(* Logix 5000 project; controller TFF vendor 1 type 14 code 107 rev 34.11; software revision 34.03; part 18 of 36 *)
(* tags used below, declared in another part *)
   AlarmControl : AlarmControl;   // Alarm Control
   ControlLoop : ControlLoop[20];   // Control Loop Array
   ControlLoop_PCV001_5ms : ALIAS FOR ControlLoop[4];   // PCV001 Control Loop
   ControlLoop_PCV101 : ALIAS FOR ControlLoop[5];   // PCV101 Control Loop
   ControlLoop_PCV101_5ms : ALIAS FOR ControlLoop[6];   // PCV101 Control Loop
   ControlLoop_PCV101Alarm : ALIAS FOR AlarmDeviation[5];   // PCV101 Control Loop Deviation Alarm
   CPU_Scanning : BOOL;   // System Scanning Flag
   DigitalOutput : BOOL[256];   // Digital Output Array these bits are sent to output cards.
   FI101 : ALIAS FOR AnalogPoint[2];   // Filtrate Flow
   FirstScanComplete : BOOL;   // First Scan Complete Flag
   LI001 : ALIAS FOR AnalogPoint[44];   // Feed Bag Volume
   Membrane_Data : Membrane_Data;   // Membrane Data
   Options : Options;   // Options List
   PCV001 : ALIAS FOR AnalogPoint[3];   // Retentate Pressure Control Valve Position
   PCV101 : ALIAS FOR AnalogPoint[4];   // Filtrate Pressure Control Valve Position
   PCV101_AO : ALIAS FOR AnalogOutput[1];   // FiltratePressure Control Valve Setpoint
   PCV101_Control : PCV_Control;   // PCV101 Control UDT
   Phase0 : ALIAS FOR Phase[0];   // Phase 0
   PLCFault : FaultRecordType;   // PLC Major Fault Record
   Rack_Murr_Node1_TF2S : IO_Station;   // Status of Node 1 TF2S
   Rack_Murr_Node1_TF3S : IO_Station;   // Status of Node 1 TF3S
   Rack_Murr_Node6_IND331_WI001 : IO_Station;   // Status of Node 6 IND331 WI001
   Rack_Murr_Node7_IND131_WI101 : IO_Station;   // Status of Node 7 IND131 WI101
   RawAnalogInputArray : INT[50];   // Array of analog input raw
   ScaleFiltering : ScaleFiltering;   // Data for Scale Filtering
   SIC001 : ALIAS FOR Drive[1];   // Feed Pump
   SIC002 : ALIAS FOR Drive[2];   // Transfer Pump
   SysControl : SysControl;   // General system status and command
   ThisSystem : SystemType;
   TMP : ALIAS FOR AnalogPoint[41];   // Trans-membrane Pressure
   Valve : Valve[100];   // Valve Array
   ValveControl : ValveControl;   // Valve Control
   WI001 : ALIAS FOR AnalogPoint[15];   // Feed Bag Weight
   WI001Alarm : ALIAS FOR AlarmAnalog[15];   // Feed Bag Weight Alarm
   WI101 : ALIAS FOR AnalogPoint[0];   // Filtrate Weight
   WI101Alarm : ALIAS FOR AlarmAnalog[0];   // Filtrate Weight Alarm
   WI102 : ALIAS FOR AnalogPoint[1];   // Customer Filtrate Weight
   WI102Alarm : ALIAS FOR AlarmAnalog[1];   // Customer Filtrate Weight Alarm
   YA10 : ALIAS FOR DigitalPoint[59];   // PLC Program Major Fault
(* MainProgram5ms, continued *)

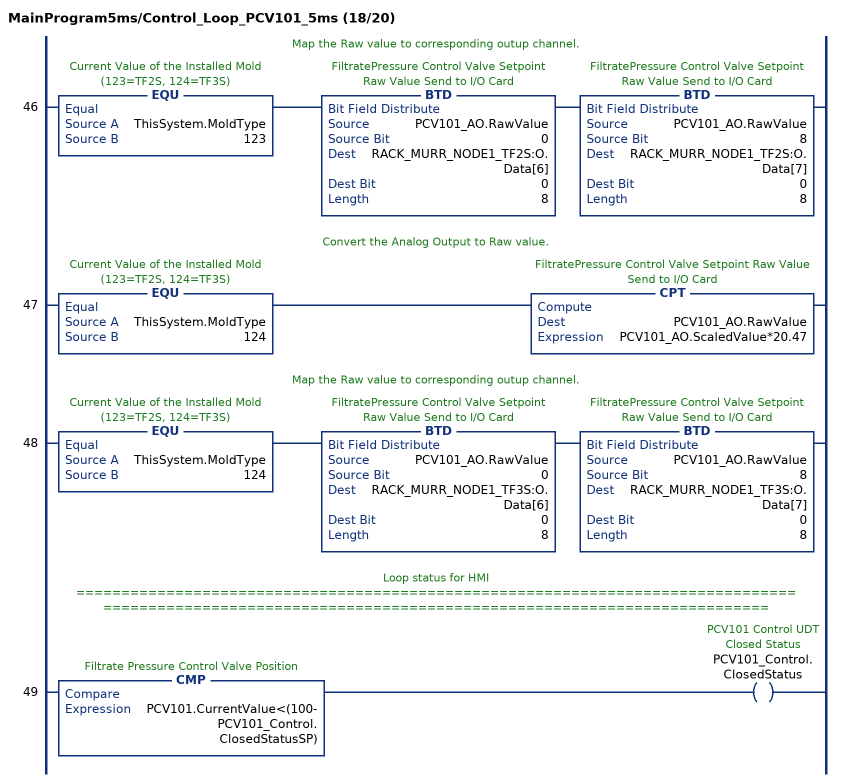
   // Map the Raw value to corresponding outup channel.
   46: EQU(ThisSystem.MoldType,123)BTD(PCV101_AO.RawValue,0,RACK_MURR_NODE1_TF2S:O.Data[6],0,8)BTD(PCV101_AO.RawValue,8,RACK_MURR_NODE1_TF2S:O.Data[7],0,8);
   // Convert the Analog Output to Raw value.
   47: EQU(ThisSystem.MoldType,124)CPT(PCV101_AO.RawValue,PCV101_AO.ScaledValue*20.47);
   // Map the Raw value to corresponding outup channel.
   48: EQU(ThisSystem.MoldType,124)BTD(PCV101_AO.RawValue,0,RACK_MURR_NODE1_TF3S:O.Data[6],0,8)BTD(PCV101_AO.RawValue,8,RACK_MURR_NODE1_TF3S:O.Data[7],0,8);
   // Loop status for HMI
   // ==========================================================================================================================================================
   49: CMP(PCV101.CurrentValue<(100-PCV101_Control.ClosedStatusSP))OTE(PCV101_Control.ClosedStatus);
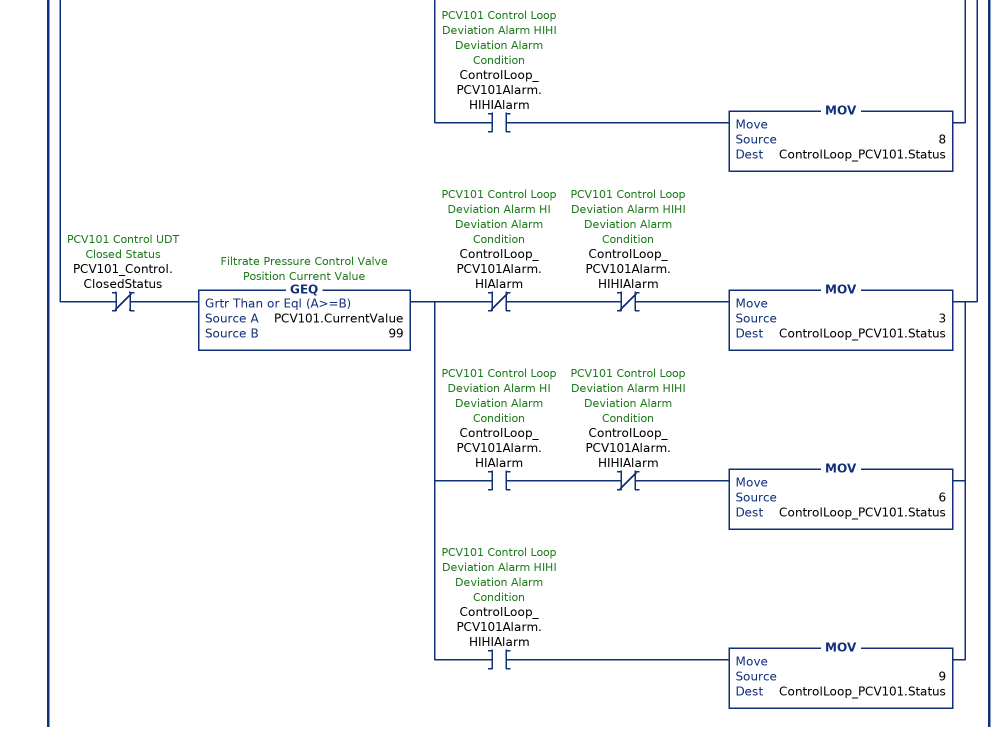
   // ControlLoop Status : 1 = PCV Close
   // ControlLoop Status : 2 = PCV Open
   // ControlLoop Status : 3 = PCV Full Open
   // ControlLoop Status : 4 = PCV Close and Non Critical alam
   // ControlLoop Status : 5 = PCV Open and Non Critical alam
   // ControlLoop Status : 6 = PCV Full Open and Non Critical alam
   // ControlLoop Status : 7 = PCV Close and Critical alam
   // ControlLoop Status : 8 = PCV Open and Critical alam
   // ControlLoop Status : 9 = PCV Full Open and Critical alam
   50: [XIC(PCV101_Control.ClosedStatus) [XIO(ControlLoop_PCV101Alarm.HIAlarm) XIO(ControlLoop_PCV101Alarm.HIHIAlarm) MOV(1,ControlLoop_PCV101.Status) ,XIC(ControlLoop_PCV101Alarm.HIAlarm) XIO(ControlLoop_PCV101Alarm.HIHIAlarm) MOV(4,ControlLoop_PCV101.Status) ,XIC(ControlLoop_PCV101Alarm.HIHIAlarm) MOV(7,ControlLoop_PCV101.Status) ] ,XIO(PCV101_Control.ClosedStatus) LES(PCV101.CurrentValue,99) [XIO(ControlLoop_PCV101Alarm.HIAlarm) XIO(ControlLoop_PCV101Alarm.HIHIAlarm) MOV(2,ControlLoop_PCV101.Status) ,XIC(ControlLoop_PCV101Alarm.HIAlarm) XIO(ControlLoop_PCV101Alarm.HIHIAlarm) MOV(5,ControlLoop_PCV101.Status) ,XIC(ControlLoop_PCV101Alarm.HIHIAlarm) MOV(8,ControlLoop_PCV101.Status) ] ,XIO(PCV101_Control.ClosedStatus) GEQ(PCV101.CurrentValue,99) [XIO(ControlLoop_PCV101Alarm.HIAlarm) XIO(ControlLoop_PCV101Alarm.HIHIAlarm) MOV(3,ControlLoop_PCV101.Status) ,XIC(ControlLoop_PCV101Alarm.HIAlarm) XIO(ControlLoop_PCV101Alarm.HIHIAlarm) MOV(6,ControlLoop_PCV101.Status) ,XIC(ControlLoop_PCV101Alarm.HIHIAlarm) MOV(9,ControlLoop_PCV101.Status) ] ];
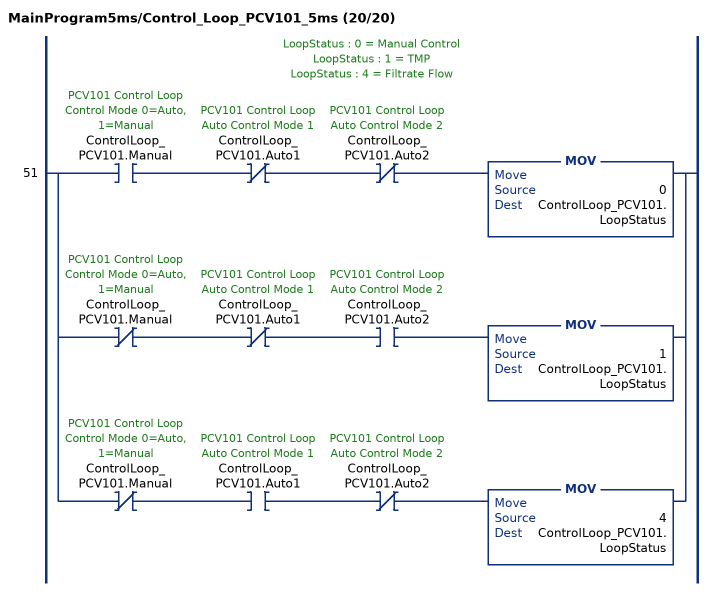
   // LoopStatus : 0 = Manual Control
   //  LoopStatus : 1 = TMP
   //  LoopStatus : 4 = Filtrate Flow
   51: [XIC(ControlLoop_PCV101.Manual) XIO(ControlLoop_PCV101.Auto1) XIO(ControlLoop_PCV101.Auto2) MOV(0,ControlLoop_PCV101.LoopStatus) ,XIO(ControlLoop_PCV101.Manual) XIO(ControlLoop_PCV101.Auto1) XIC(ControlLoop_PCV101.Auto2) MOV(1,ControlLoop_PCV101.LoopStatus) ,XIO(ControlLoop_PCV101.Manual) XIC(ControlLoop_PCV101.Auto1) XIO(ControlLoop_PCV101.Auto2) MOV(4,ControlLoop_PCV101.LoopStatus) ];
END_ROUTINE

ROUTINE FaultRoutine   (* ladder *)
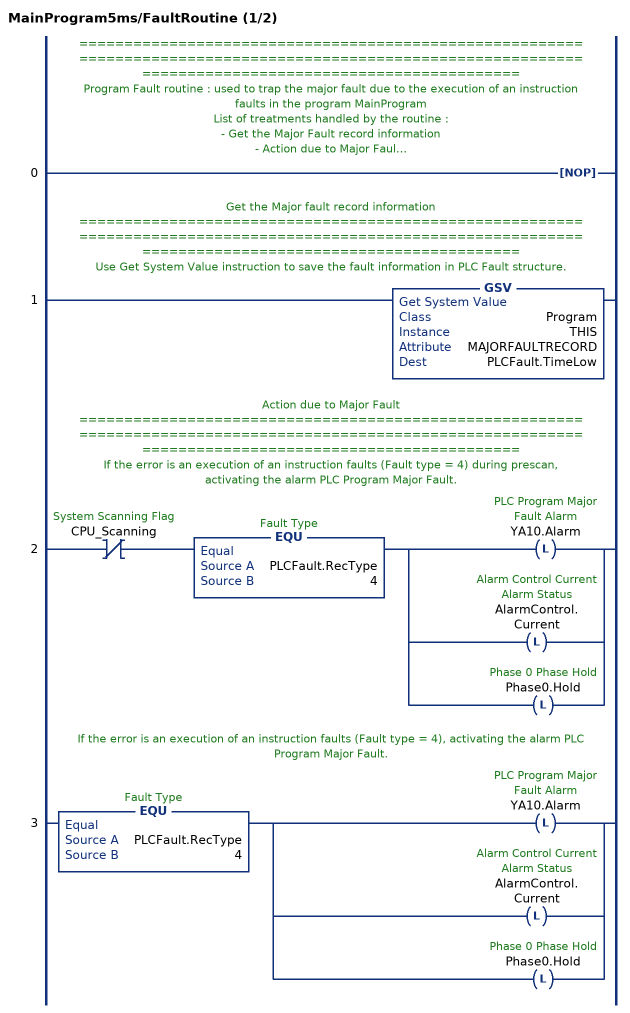
   // ==========================================================================================================================================================
   //                                                               Program Fault routine : used to trap the major fault due to the execution of an instruction faults in the program MainProgram
   //                                                     List of treatments handled by the routine :
   //                                                          - Get the Major Fault record information
   //                                                          - Action due to Major Fault
   //                                                     -----------------------------------------------------------------------------------------------------------------------------------------------------
   //                                                     History
   //                                                          2019-AUG-13 - Actemium - B. Roch - Initial version for Candidate Release 3.00.00.00.a
   // ==========================================================================================================================================================
   0: NOP();
   // Get the Major fault record information
   // ==========================================================================================================================================================
   // Use Get System Value instruction to save the fault information in PLC Fault structure.
   1: GSV(Program,THIS,MAJORFAULTRECORD,PLCFault.TimeLow);
   // Action due to Major Fault
   // ==========================================================================================================================================================
   // If the error is an execution of an instruction faults (Fault type = 4) during prescan, activating the alarm PLC Program Major Fault.
   2: XIO(CPU_Scanning)EQU(PLCFault.RecType,4)[OTL(YA10.Alarm) ,OTL(AlarmControl.Current) ,OTL(Phase0.Hold) ];
   // If the error is an execution of an instruction faults (Fault type = 4), activating the alarm PLC Program Major Fault.
   3: EQU(PLCFault.RecType,4)[OTL(YA10.Alarm) ,OTL(AlarmControl.Current) ,OTL(Phase0.Hold) ];
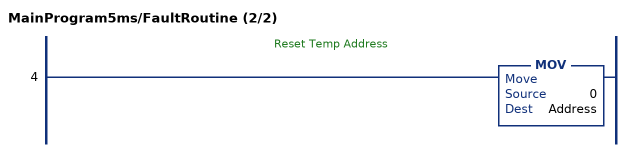
   // Reset Temp Address
   4: MOV(0,Address);
END_ROUTINE

ROUTINE Input_Analog_HighSpeed   (* ladder *)
// HighSpeed Analog Input Scaling
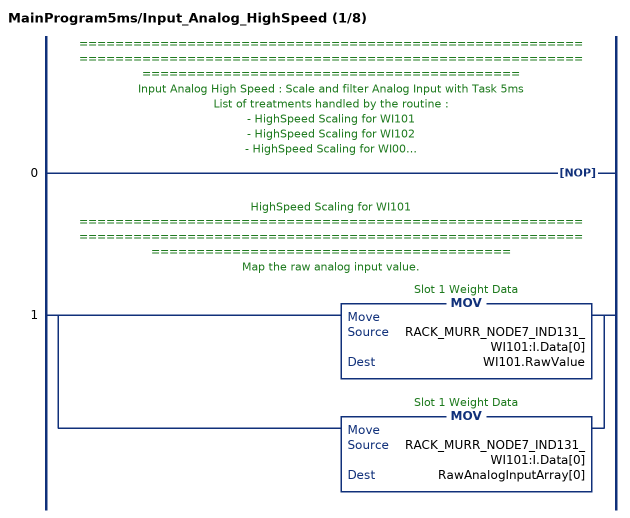
   // ==========================================================================================================================================================
   //                                                  Input Analog High Speed : Scale and filter Analog Input with Task 5ms
   //                                                     List of treatments handled by the routine :
   //                                                     - HighSpeed Scaling for WI101
   //                                                     - HighSpeed Scaling for WI102
   //                                                     - HighSpeed Scaling for WI001
   //                                                     - Scale Filtering processing
   //                                                     - Alarm Process Value Initialization
   //                                                     -----------------------------------------------------------------------------------------------------------------------------------------------------
   //                                                     History
   //                                                   2019-AUG-13 - Actemium - B. Roch - Initial version for Candidate Release 3.00.00.00.a                    		2019-SEP-11 - ACTEMIUM - Q. Spindler - Modifications for Candidate Release 3.00.00.00.c
   // 					- Change raw value for WI102 to 1
   // ==========================================================================================================================================================
   0: NOP();
   // HighSpeed Scaling for WI101
   // ========================================================================================================================================================
   // Map the raw analog input value.
   1: [MOV(RACK_MURR_NODE7_IND131_WI101:I.Data[0],WI101.RawValue) ,MOV(RACK_MURR_NODE7_IND131_WI101:I.Data[0],RawAnalogInputArray[0]) ];
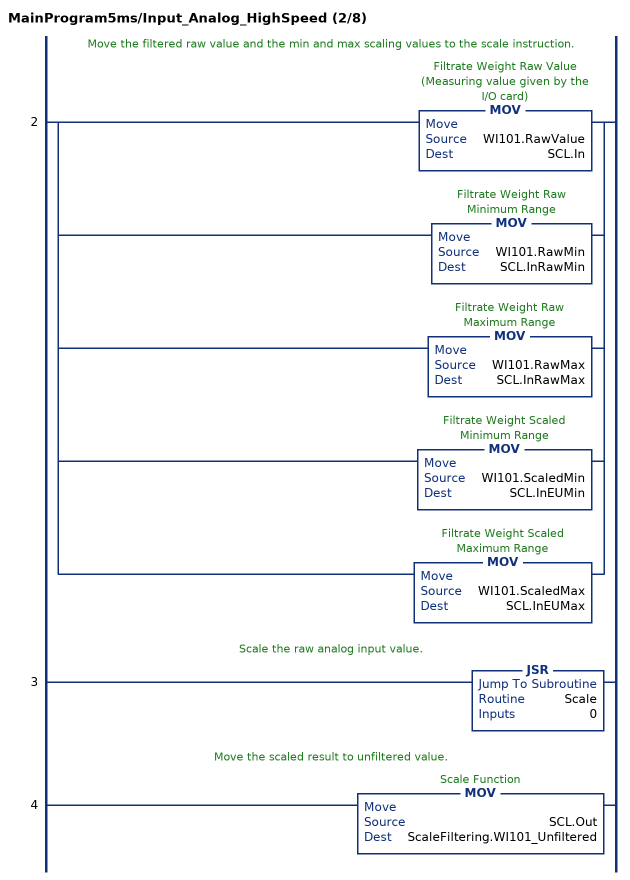
   // Move the filtered raw value and the min and max scaling values to the scale instruction.
   2: [MOV(WI101.RawValue,SCL.In) ,MOV(WI101.RawMin,SCL.InRawMin) ,MOV(WI101.RawMax,SCL.InRawMax) ,MOV(WI101.ScaledMin,SCL.InEUMin) ,MOV(WI101.ScaledMax,SCL.InEUMax) ];
   // Scale the raw analog input value.
   3: JSR(Scale,0);
   // Move the scaled result to unfiltered value.
   4: MOV(SCL.Out,ScaleFiltering.WI101_Unfiltered);
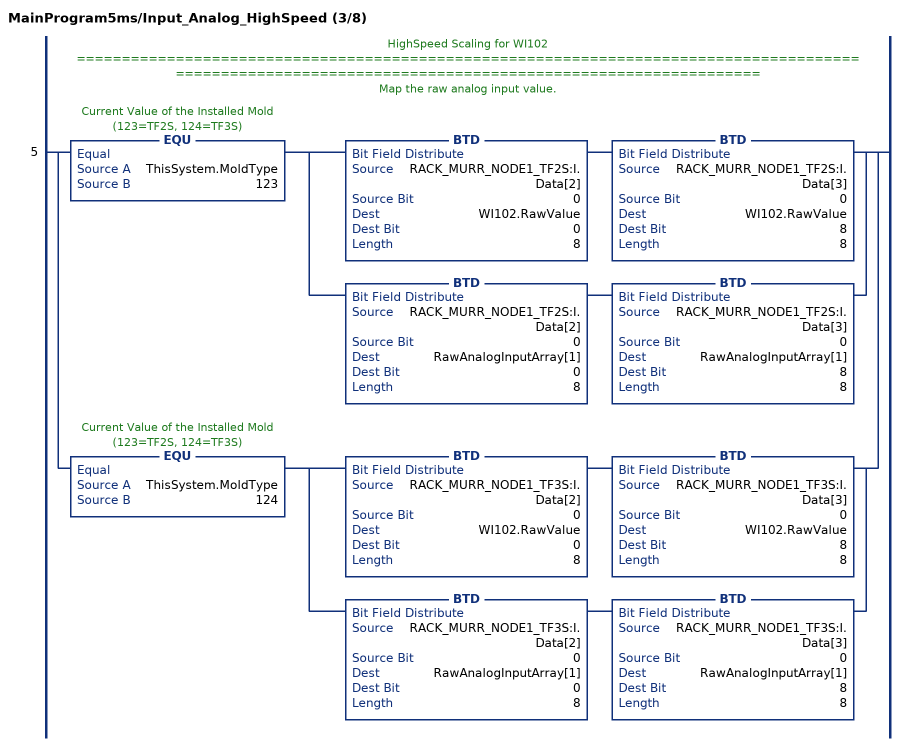
   // HighSpeed Scaling for WI102
   // ========================================================================================================================================================
   // Map the raw analog input value.
   5: [EQU(ThisSystem.MoldType,123) [BTD(RACK_MURR_NODE1_TF2S:I.Data[2],0,WI102.RawValue,0,8) BTD(RACK_MURR_NODE1_TF2S:I.Data[3],0,WI102.RawValue,8,8) ,BTD(RACK_MURR_NODE1_TF2S:I.Data[2],0,RawAnalogInputArray[1],0,8) BTD(RACK_MURR_NODE1_TF2S:I.Data[3],0,RawAnalogInputArray[1],8,8) ] ,EQU(ThisSystem.MoldType,124) [BTD(RACK_MURR_NODE1_TF3S:I.Data[2],0,WI102.RawValue,0,8) BTD(RACK_MURR_NODE1_TF3S:I.Data[3],0,WI102.RawValue,8,8) ,BTD(RACK_MURR_NODE1_TF3S:I.Data[2],0,RawAnalogInputArray[1],0,8) BTD(RACK_MURR_NODE1_TF3S:I.Data[3],0,RawAnalogInputArray[1],8,8) ] ];
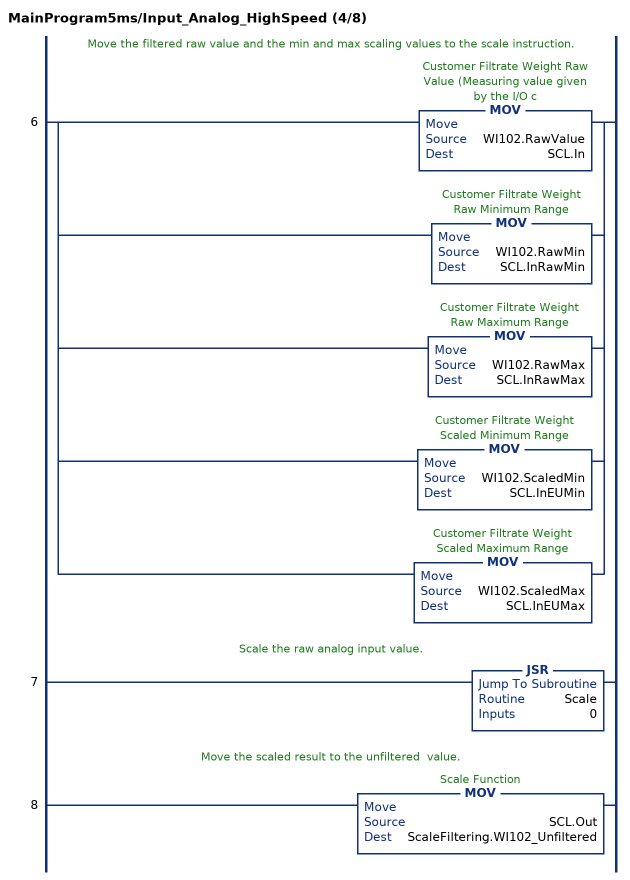
   // Move the filtered raw value and the min and max scaling values to the scale instruction.
   6: [MOV(WI102.RawValue,SCL.In) ,MOV(WI102.RawMin,SCL.InRawMin) ,MOV(WI102.RawMax,SCL.InRawMax) ,MOV(WI102.ScaledMin,SCL.InEUMin) ,MOV(WI102.ScaledMax,SCL.InEUMax) ];
   // Scale the raw analog input value.
   7: JSR(Scale,0);
   // Move the scaled result to the unfiltered  value.
   8: MOV(SCL.Out,ScaleFiltering.WI102_Unfiltered);
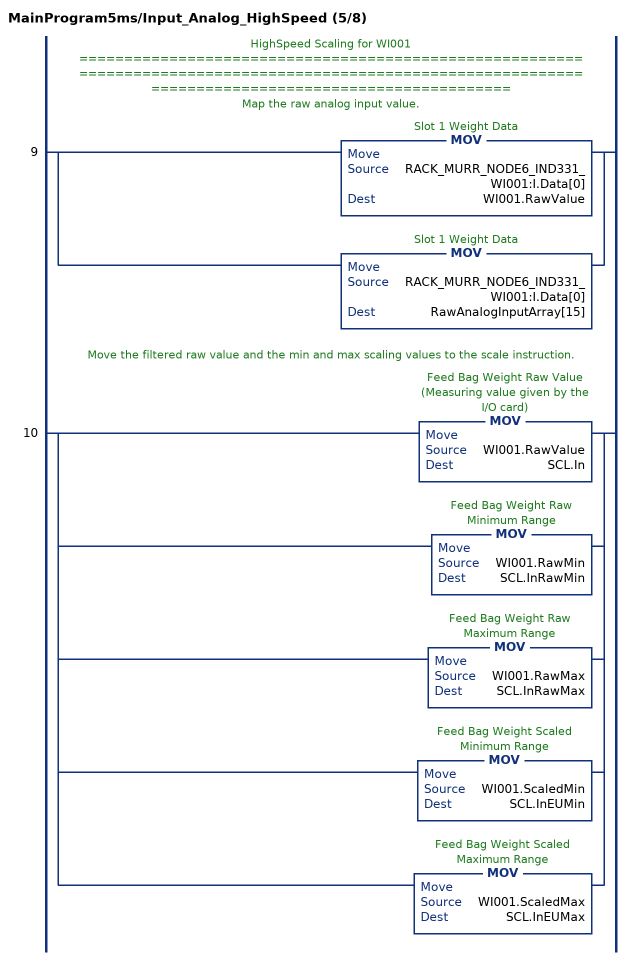
   // HighSpeed Scaling for WI001
   // ========================================================================================================================================================
   // Map the raw analog input value.
   9: [MOV(RACK_MURR_NODE6_IND331_WI001:I.Data[0],WI001.RawValue) ,MOV(RACK_MURR_NODE6_IND331_WI001:I.Data[0],RawAnalogInputArray[15]) ];
   // Move the filtered raw value and the min and max scaling values to the scale instruction.
   10: [MOV(WI001.RawValue,SCL.In) ,MOV(WI001.RawMin,SCL.InRawMin) ,MOV(WI001.RawMax,SCL.InRawMax) ,MOV(WI001.ScaledMin,SCL.InEUMin) ,MOV(WI001.ScaledMax,SCL.InEUMax) ];
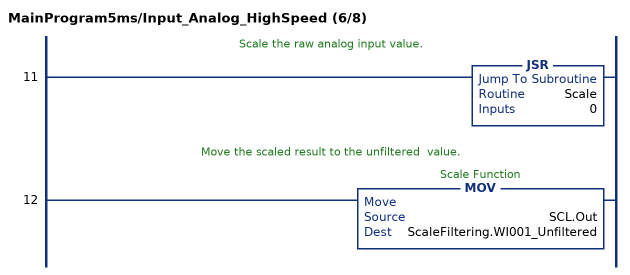
   // Scale the raw analog input value.
   11: JSR(Scale,0);
   // Move the scaled result to the unfiltered  value.
   12: MOV(SCL.Out,ScaleFiltering.WI001_Unfiltered);
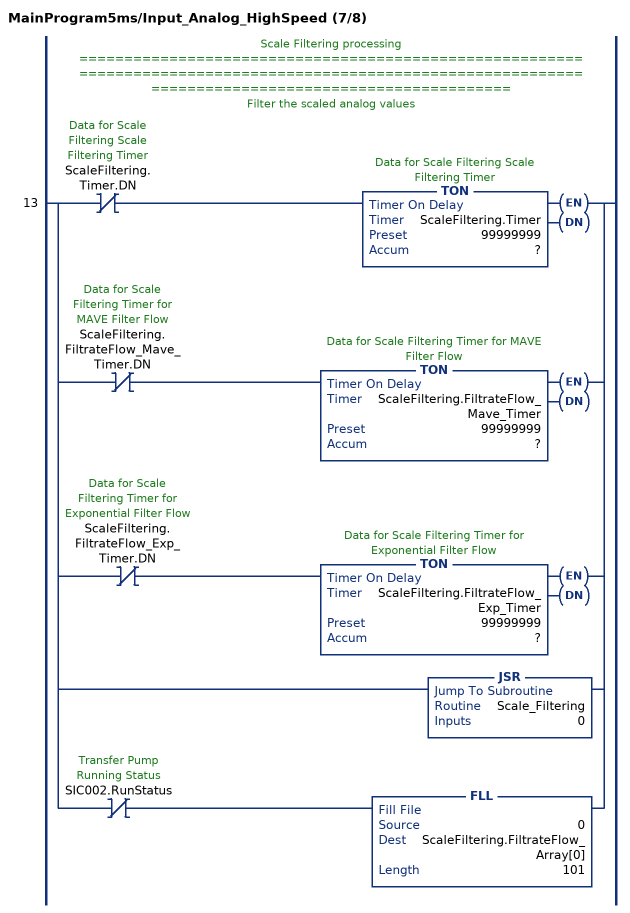
   // Scale Filtering processing
   // ========================================================================================================================================================
   // Filter the scaled analog values
   13: [XIO(ScaleFiltering.Timer.DN) TON(ScaleFiltering.Timer,?,?) ,XIO(ScaleFiltering.FiltrateFlow_Mave_Timer.DN) TON(ScaleFiltering.FiltrateFlow_Mave_Timer,?,?) ,XIO(ScaleFiltering.FiltrateFlow_Exp_Timer.DN) TON(ScaleFiltering.FiltrateFlow_Exp_Timer,?,?) ,JSR(Scale_Filtering,0) ,XIO(SIC002.RunStatus) FLL(0,ScaleFiltering.FiltrateFlow_Array[0],101) ];
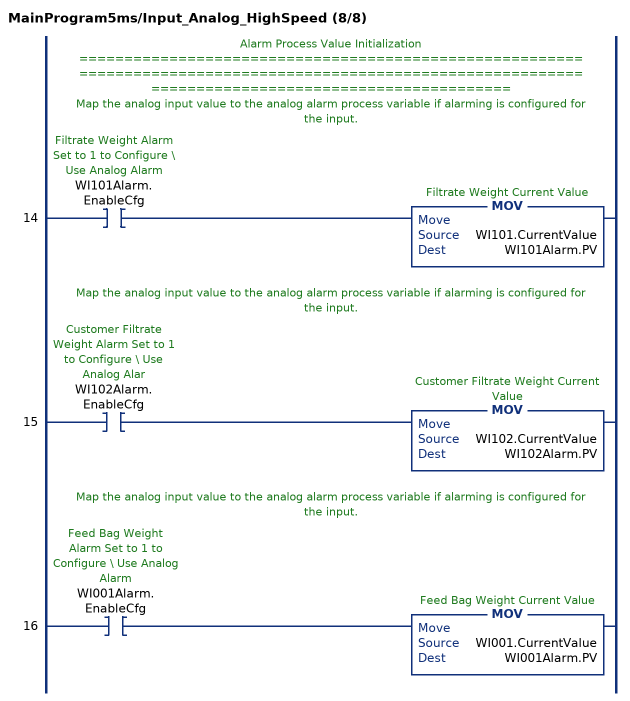
   // Alarm Process Value Initialization
   // ========================================================================================================================================================
   // Map the analog input value to the analog alarm process variable if alarming is configured for the input.
   14: XIC(WI101Alarm.EnableCfg)MOV(WI101.CurrentValue,WI101Alarm.PV);
   // Map the analog input value to the analog alarm process variable if alarming is configured for the input.
   15: XIC(WI102Alarm.EnableCfg)MOV(WI102.CurrentValue,WI102Alarm.PV);
   // Map the analog input value to the analog alarm process variable if alarming is configured for the input.
   16: XIC(WI001Alarm.EnableCfg)MOV(WI001.CurrentValue,WI001Alarm.PV);
END_ROUTINE

ROUTINE MainRoutine   (* ladder *)
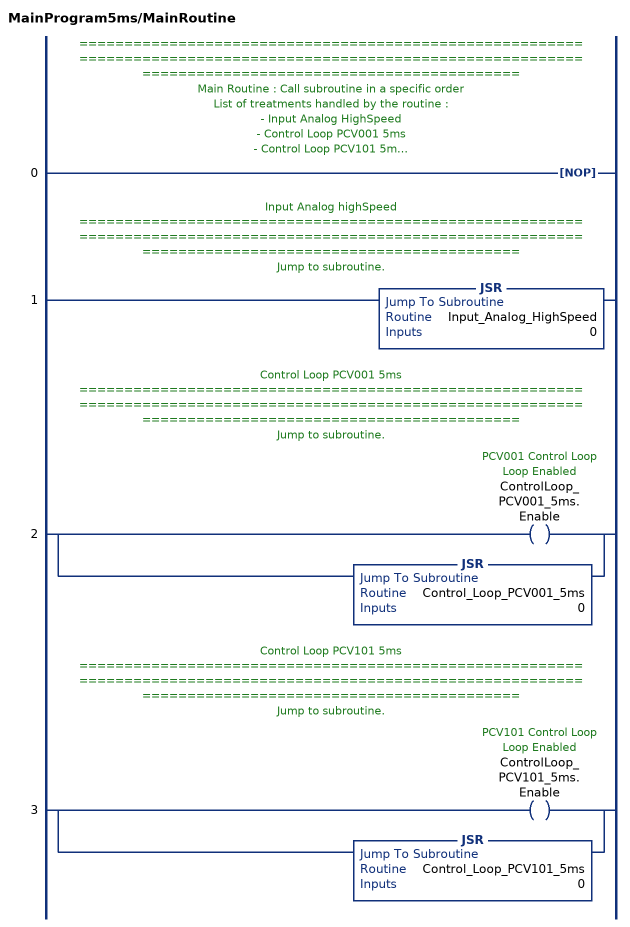
   // ==========================================================================================================================================================
   //                                                  Main Routine : Call subroutine in a specific order
   //                                                     List of treatments handled by the routine :
   //                                                - Input Analog HighSpeed
   //                                                - Control Loop PCV001 5ms
   //                                                - Control Loop PCV101 5ms
   //                                                     -----------------------------------------------------------------------------------------------------------------------------------------------------
   //                                                     History
   //                                                        2019-AUG-13 - Actemium - B. Roch - Initial version for Candidate Release 3.00.00.00.a
   // ==========================================================================================================================================================
   0: NOP();
   // Input Analog highSpeed
   // ==========================================================================================================================================================
   // Jump to subroutine.
   1: JSR(Input_Analog_HighSpeed,0);
   // Control Loop PCV001 5ms
   // ==========================================================================================================================================================
   // Jump to subroutine.
   2: [OTE(ControlLoop_PCV001_5ms.Enable) ,JSR(Control_Loop_PCV001_5ms,0) ];
   // Control Loop PCV101 5ms
   // ==========================================================================================================================================================
   // Jump to subroutine.
   3: [OTE(ControlLoop_PCV101_5ms.Enable) ,JSR(Control_Loop_PCV101_5ms,0) ];
END_ROUTINE

ROUTINE Scale   (* function block diagram *)
// Scale Routine
   SHEET 1
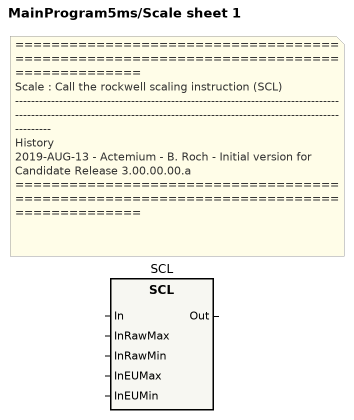
   // ======================================================================================
   // Scale : Call the rockwell scaling instruction (SCL)
   // ------------------------------------------------------------------------------------------------------------------------------------------------------------------
   // ---------
   // History
   //    2019-AUG-13 - Actemium - B. Roch - Initial version for Candidate Release 3.00.00.00.a
   // ======================================================================================
   SCL : SCL();   // unwired pins: In InRawMax InRawMin InEUMax InEUMin Out
END_ROUTINE

ROUTINE Scale_Filtering   (* structured text *)
   
   (* =======================================================================
   	Scale Filtering : calculations of Filtered value
   
   	List of treatments
   		- Initialize Volume
   		- WI001 Feed Bag Volume Calculation
   		- Moving Average Filtering for Filtrate Volume
   		- Moving Average Filtering for Filtrate Flow
   		- Exponential Filtering for Filtrate Volume
   		- Exponential Filtering for Filtrate Flow
   		- Analog Input processing
   
   -----------------------------------------------------------------------------------------------------------------------------------------------------
   	History
   		2019-AUG-13 - ACTEMIUM - B. Roch - Initial version for Candidate Release 3.00.00.00.a
   		2019-SEP-17 - ACTEMIUM - Q. Spindler - Modifications for Candidate Release 3.00.00.00.c
   					- Bypass CurrentValue calculation when in simulation mode
   					- Remove Initialize Values as they will be stored in CCPSettings
   =============================================================================================================================*)
   
   
   
   (* Initialize Volume
   =============================================================================================================================*)
   
   // Compute Volume values based on Unfiltered Weight and Density
   ScaleFiltering.FeedBagVolume := ScaleFiltering.WI001_Unfiltered / Membrane_Data.Density;
   ScaleFiltering.FiltrateVolume101 := ScaleFiltering.WI101_Unfiltered / Membrane_Data.Density;
   ScaleFiltering.FiltrateVolume102 := ScaleFiltering.WI102_Unfiltered / Membrane_Data.Density;
   
   
   //Check that the minimum sample rate have met
   If ScaleFiltering.Timer.ACC > ScaleFiltering.Sample_Rate Then
   
   (* WI001 Feed Bag Volume Calculation
   =============================================================================================================================*)
   
   		//Compute the feed bag volume and Weight using the moving average filter
   		ScaleFiltering.FeedBagVolume_MAVE.In := ScaleFiltering.FeedBagVolume;
   		MAVE(ScaleFiltering.FeedBagVolume_MAVE, ScaleFiltering.FeedBagVolume_Array);
   		If Not SysControl.Simulate Then
   			LI001.CurrentValue := ScaleFiltering.FeedBagVolume_MAVE.Out;
   			WI001.CurrentValue := ScaleFiltering.FeedBagVolume_MAVE.Out * Membrane_Data.Density;
   		Else
   			LI001.CurrentValue := WI001.CurrentValue / Membrane_Data.Density;
   		End_If;
   
   (* Moving Average Filtering for Filtrate Volume
   =============================================================================================================================*)
   
   		//Compute the Filtrate volume and Weight (Merck) using the moving average filter
   		ScaleFiltering.FiltrateVolume101_MAVE.In := ScaleFiltering.FiltrateVolume101;
   		MAVE(ScaleFiltering.FiltrateVolume101_MAVE, ScaleFiltering.FiltrateVolume101_Array);
   		ScaleFiltering.FiltrateVolume101_MaveFiltered := ScaleFiltering.FiltrateVolume101_MAVE.Out;
   		ScaleFiltering.Weight101_MaveFiltered := ScaleFiltering.FiltrateVolume101_MAVE.Out * Membrane_Data.Density;
   
   		//Compute the Filtrate volume and Weight (Customer) using the moving average filter
   		ScaleFiltering.FiltrateVolume102_MAVE.In := ScaleFiltering.FiltrateVolume102;
   		MAVE(ScaleFiltering.FiltrateVolume102_MAVE, ScaleFiltering.FiltrateVolume102_Array);
   		ScaleFiltering.FiltrateVolume102_MaveFiltered := ScaleFiltering.FiltrateVolume102_MAVE.Out;
   		ScaleFiltering.Weight102_MaveFiltered := ScaleFiltering.FiltrateVolume102_MAVE.Out * Membrane_Data.Density;
   
   		//Set the Filtered Volume based on current options configuration
   		If Options.WI101 Then;
   			ScaleFiltering.FiltrateVolume_MaveFiltered := ScaleFiltering.FiltrateVolume101_MaveFiltered;
   		ElsIf Options.WI102 Then;
   			ScaleFiltering.FiltrateVolume_MaveFiltered := ScaleFiltering.FiltrateVolume102_MaveFiltered;
   		End_If;
   
   (* Moving Average Filtering for Filtrate Flow
   =============================================================================================================================*)
   
   		If SIC001.RunStatus Then
   			If (ScaleFiltering.FiltrateFlow_Mave_Timer.ACC > ScaleFiltering.FiltrateFlow_Mave_Sample_Rate) Then
   				If (ABS(ScaleFiltering.FiltrateVolume_MaveFiltered - ScaleFiltering.FiltrateVolume_MaveFiltered_Prev) >= 0.01) Then
   					//Compute the Filtrate Flow rate
   					//Filtrate Flow Rate = ((Current Volume - Previous Volume) / Time Elapsed (in s)) * 60
   					ScaleFiltering.FiltrateFlow := ((ScaleFiltering.FiltrateVolume_MaveFiltered - ScaleFiltering.FiltrateVolume_MaveFiltered_Prev) / (ScaleFiltering.FiltrateFlow_Mave_Timer.ACC / 1000))*60;
   					ScaleFiltering.FiltrateVolume_MaveFiltered_Prev := ScaleFiltering.FiltrateVolume_MaveFiltered;
   
   					//Compute the Filtrate Flow Rate using the moving average filter
   					ScaleFiltering.FiltrateFlow_MAVE.In := ScaleFiltering.FiltrateFlow;
   					MAVE(ScaleFiltering.FiltrateFlow_MAVE, ScaleFiltering.FiltrateFlow_Array);
   					ScaleFiltering.FiltrateFlow_MaveFiltered := ScaleFiltering.FiltrateFlow_MAVE.Out;
   
   					ScaleFiltering.FiltrateFlow_Mave_Timer.ACC :=0;
   				End_If;
   			End_If;
   		Else
   			ScaleFiltering.FiltrateFlow_MaveFiltered := 0;
   			ScaleFiltering.FiltrateFlow_Mave_Timer.ACC :=0;
   		End_If;
   
   (* Exponential Filtering for Filtrate Volume
   =============================================================================================================================*)
   
   	//Compute the Filtrate volume using the Exponential filter
   	ScaleFiltering.FiltrateVolume101_ExpFiltered := (ScaleFiltering.FiltrateVolume101_ExpConst * ScaleFiltering.FiltrateVolume101_ExpFiltered) + ((1-ScaleFiltering.FiltrateVolume101_ExpConst)*ScaleFiltering.FiltrateVolume101);
   	ScaleFiltering.FiltrateVolume102_ExpFiltered := (ScaleFiltering.FiltrateVolume102_ExpConst * ScaleFiltering.FiltrateVolume102_ExpFiltered) + ((1-ScaleFiltering.FiltrateVolume102_ExpConst)*ScaleFiltering.FiltrateVolume102);
   
   	//Compute the Filtrate Weight using the filtered volume and density parameter
   	ScaleFiltering.Weight101_ExpFiltered := ScaleFiltering.FiltrateVolume101_ExpFiltered * Membrane_Data.Density;
   	ScaleFiltering.Weight102_ExpFiltered := ScaleFiltering.FiltrateVolume102_ExpFiltered * Membrane_Data.Density;
   
   	//Set the Filtered Volume based on current options configuration
   	If Options.WI101 Then;
   		ScaleFiltering.FiltrateVolume_ExpFiltered := ScaleFiltering.FiltrateVolume101_ExpFiltered;
   	ElsIf Options.WI102 Then;
   		ScaleFiltering.FiltrateVolume_ExpFiltered := ScaleFiltering.FiltrateVolume102_ExpFiltered;
   	End_If;
   
   (* Exponential Filtering for Filtrate Flow
   =============================================================================================================================*)
   
   	//Compute the Filtrate Flow rate
   	If ScaleFiltering.FiltrateFlow_Exp_Timer.ACC > ScaleFiltering.FiltrateFlow_Exp_Sample_Rate Then
   		ScaleFiltering.FiltrateFlow := ((ScaleFiltering.FiltrateVolume_ExpFiltered - ScaleFiltering.FiltrateVolume_ExpFiltered_Prev) / (ScaleFiltering.FiltrateFlow_Exp_Timer.ACC / 1000))*60;
   		ScaleFiltering.FiltrateVolume_ExpFiltered_Prev := ScaleFiltering.FiltrateVolume_ExpFiltered;
   
   		ScaleFiltering.FiltrateFlow_ExpFiltered := (ScaleFiltering.FiltrateFlow_ExpConst * ScaleFiltering.FiltrateFlow_ExpFiltered) + ((1-ScaleFiltering.FiltrateFlow_ExpConst) * ScaleFiltering.FiltrateFlow);
   		ScaleFiltering.FiltrateFlow_Exp_Timer.ACC := 0;
   	End_If;
   
   
   
   (* Analog Input processing
   =============================================================================================================================*)
   	//Assign Value to corresponding input
   	//Populate Analog Inputs when Pump is running and FI101 is calculated value
   	If SIC001.RunStatus AND (NOT FI101.RealCfg) Then
   		//No Filtering
   		If ScaleFiltering.CurrentFilter = 0 Then
   			If Not SysControl.Simulate Then
   				WI101.CurrentValue := ScaleFiltering.FiltrateVolume101 * Membrane_Data.Density;
   				WI102.CurrentValue := ScaleFiltering.FiltrateVolume102 * Membrane_Data.Density;
   				FI101.CurrentValue := ((ScaleFiltering.FiltrateVolume101 - ScaleFiltering.FiltrateVolume101_Filtered_Prev) / (ScaleFiltering.Timer.ACC / 1000))*60;
   			End_if;
   			ScaleFiltering.FiltrateVolume101_Filtered_Prev := ScaleFiltering.FiltrateVolume101;
   		End_If;
   
   		//Moving Average Filter Active
   		If ScaleFiltering.CurrentFilter = 1 Then
   			If Not SysControl.Simulate Then
   				WI101.CurrentValue := ScaleFiltering.Weight101_MaveFiltered;
   				WI102.CurrentValue := ScaleFiltering.Weight102_MaveFiltered;
   				FI101.CurrentValue := ScaleFiltering.FiltrateFlow_MaveFiltered;
   			End_If;
   		End_If;
   
   		//Exponential Linear Recursive Filter active
   		If ScaleFiltering.CurrentFilter = 2 Then
   			If Not SysControl.Simulate Then
   				WI101.CurrentValue := ScaleFiltering.Weight101_ExpFiltered;
   				WI102.CurrentValue := ScaleFiltering.Weight102_ExpFiltered;
   				FI101.CurrentValue := ScaleFiltering.FiltrateFlow_ExpFiltered;
   			End_If;
   		End_If;
   
   	Else //On
   		// Only populate with 0.00 when FI101 is a calculated value and the Feed Pump is OFF
   		If NOT FI101.RealCfg Then
   			If Not SysControl.Simulate Then
   				FI101.CurrentValue := 0.00;
   			End_If;
   		End_If;
   
   		If ScaleFiltering.CurrentFilter = 0 Then //No Filtering
   			If Not SysControl.Simulate Then
   				WI101.CurrentValue := ScaleFiltering.FiltrateVolume101 * Membrane_Data.Density;
   				WI102.CurrentValue := ScaleFiltering.FiltrateVolume102 * Membrane_Data.Density;
   			End_If;
   		End_If;
   
   		If ScaleFiltering.CurrentFilter = 1 Then //Moving Average Filter Active
   			If Not SysControl.Simulate Then
   				WI101.CurrentValue := ScaleFiltering.Weight101_MaveFiltered;
   				WI102.CurrentValue := ScaleFiltering.Weight102_MaveFiltered;
   			End_If;
   		End_If;
   
   		If ScaleFiltering.CurrentFilter = 2 Then //Exponential Linear Recursive Filter active
   			If Not SysControl.Simulate Then
   				WI101.CurrentValue := ScaleFiltering.Weight101_ExpFiltered;
   				WI102.CurrentValue := ScaleFiltering.Weight102_ExpFiltered;
   			End_If;
   		End_If;
   	End_If;
   
   	ScaleFiltering.Timer.ACC := 0;
   End_If;
   
   (*Reset Filtrate value if option is active*)
   IF Options.No_Filtrate_Measurement THEN
   	FI101.CurrentValue := 0.00;
   END_IF;
END_ROUTINE
END_PROGRAM

PROGRAM Process   (* main routine MainRoutine, fault routine FaultRoutine *)
VAR
   Address : DINT;   // Temp Address
   Address2 : DINT := 41;   // Temp Address
   AddressPump1 : DINT := 1;   // Temp Address for Pump 1
   AddressPump2 : DINT := 2;   // Temp Address for Pump 2
   AlarmInhibit_Timer : TIMER := (PRE := 500, ACC := 500);
   BufferSteps0_Prev : STRING25 := '67';
   Config : Configuration := (IndexA0 := 25, IndexAP := 50, IndexDP := 150, IndexDr := 11, IndeXValve := 100, IndexCL := 20, IndexFlowpath := 61);   // Index Array used in configuration routines
   FeedBagLevel_PID_Settings : INT;   // Index
   FeedPump_PID_Settings : INT;   // Index
   Index : DINT;   // Index
   Index2 : DINT;   // Index
   Index3 : DINT;   // Index
   index4 : DINT := 21;   // Index
   NewSystem : DINT := 124;
   ON_OFF : BOOL;
   ONS_PID02 : BOOL;
   PCV001_PID_Settings : INT;
   PCV101_PID_Settings : INT;
   RecipeStepLog_DateTime_Empty : STRING25;   // Empty String
   RecipeStepLog_DateTime_Log : STRING25 := '11/08/2026 1:25:40 A';   // Last Date Time received from HMI
   RecipeStepLog_DateTime_Prev : STRING25 := '11/08/2026 1:25:40 A';
   RecipeStepLog_Timer : TIMER := (PRE := 15000, ACC := 15003, EN := 1, DN := 1);   // RecipeStepLog Watchdog Timer
   sBar1 : STRING5 := 'bar';
   sBar2 : STRING5 := 'Bar';
   sBar3 : STRING5 := 'BAR';
   SCL : SCALE := (Status := 16#0000_0003, InstructFault := 1, InRawRangeInv := 1);   // Scale Instruction
END_VAR

ROUTINE Alarm   (* ladder *)
// Alarm Routine
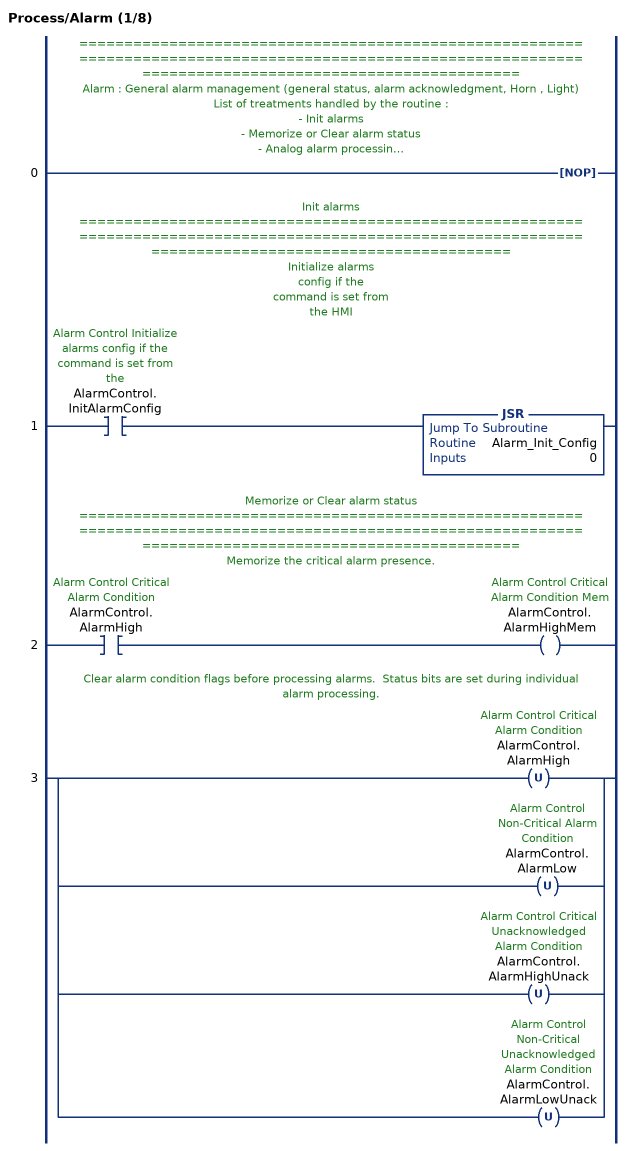
   // ==========================================================================================================================================================
   //                                                                                     Alarm : General alarm management (general status, alarm acknowledgment, Horn , Light)
   //                                                     List of treatments handled by the routine :
   //                                                         - Init alarms
   //                                                          - Memorize or Clear alarm status
   //                                                          - Analog alarm processing
   //                                                          - Deviation alarm processing
   //                                                          - Digital alarm processing
   //                                                          - General alarm status
   //                                                          - Flash control
   //                                                          - Alarm Horn
   //                                                          - Alarm Light
   //                                                          - Alarm acknowledgment
   //                                                          - Output processing
   //                                                     -----------------------------------------------------------------------------------------------------------------------------------------------------
   //                                                     History
   //                                                          2019-AUG-13 - Actemium - B. Roch - Initial version for Candidate Release 3.00.00.00.a
   //                                                           2020-Sep-28 - Merck - Q.Spindler - Modifications for Candidate Release 3.00.00.01.a
   // - Add Alarm Init Call
   // ==========================================================================================================================================================
   0: NOP();
   // Init alarms
   // ========================================================================================================================================================
   //  Initialize alarms
   // config if the
   // command is set from
   // the HMI
   1: XIC(AlarmControl.InitAlarmConfig)JSR(Alarm_Init_Config,0);
   // Memorize or Clear alarm status
   // ==========================================================================================================================================================
   // Memorize the critical alarm presence.
   2: XIC(AlarmControl.AlarmHigh)OTE(AlarmControl.AlarmHighMem);
   // Clear alarm condition flags before processing alarms.  Status bits are set during individual alarm processing.
   3: [OTU(AlarmControl.AlarmHigh) ,OTU(AlarmControl.AlarmLow) ,OTU(AlarmControl.AlarmHighUnack) ,OTU(AlarmControl.AlarmLowUnack) ];
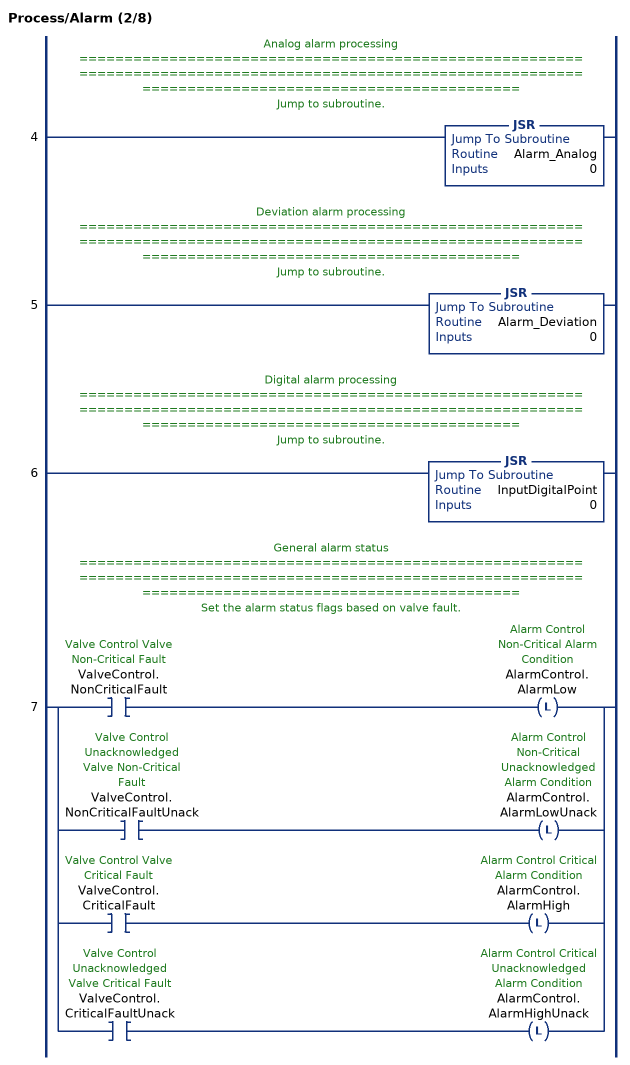
   // Analog alarm processing
   // ==========================================================================================================================================================
   // Jump to subroutine.
   4: JSR(Alarm_Analog,0);
   // Deviation alarm processing
   // ==========================================================================================================================================================
   // Jump to subroutine.
   5: JSR(Alarm_Deviation,0);
   // Digital alarm processing
   // ==========================================================================================================================================================
   // Jump to subroutine.
   6: JSR(InputDigitalPoint,0);
   // General alarm status
   // ==========================================================================================================================================================
   // Set the alarm status flags based on valve fault.
   7: [XIC(ValveControl.NonCriticalFault) OTL(AlarmControl.AlarmLow) ,XIC(ValveControl.NonCriticalFaultUnack) OTL(AlarmControl.AlarmLowUnack) ,XIC(ValveControl.CriticalFault) OTL(AlarmControl.AlarmHigh) ,XIC(ValveControl.CriticalFaultUnack) OTL(AlarmControl.AlarmHighUnack) ];
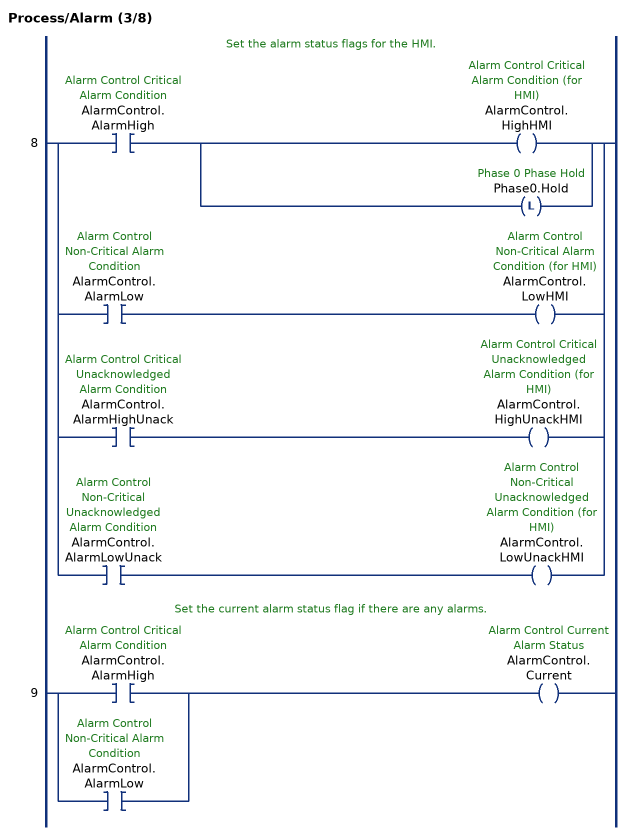
   // Set the alarm status flags for the HMI.
   8: [XIC(AlarmControl.AlarmHigh) [OTE(AlarmControl.HighHMI) ,OTL(Phase0.Hold) ] ,XIC(AlarmControl.AlarmLow) OTE(AlarmControl.LowHMI) ,XIC(AlarmControl.AlarmHighUnack) OTE(AlarmControl.HighUnackHMI) ,XIC(AlarmControl.AlarmLowUnack) OTE(AlarmControl.LowUnackHMI) ];
   // Set the current alarm status flag if there are any alarms.
   9: [XIC(AlarmControl.AlarmHigh) ,XIC(AlarmControl.AlarmLow) ]OTE(AlarmControl.Current);
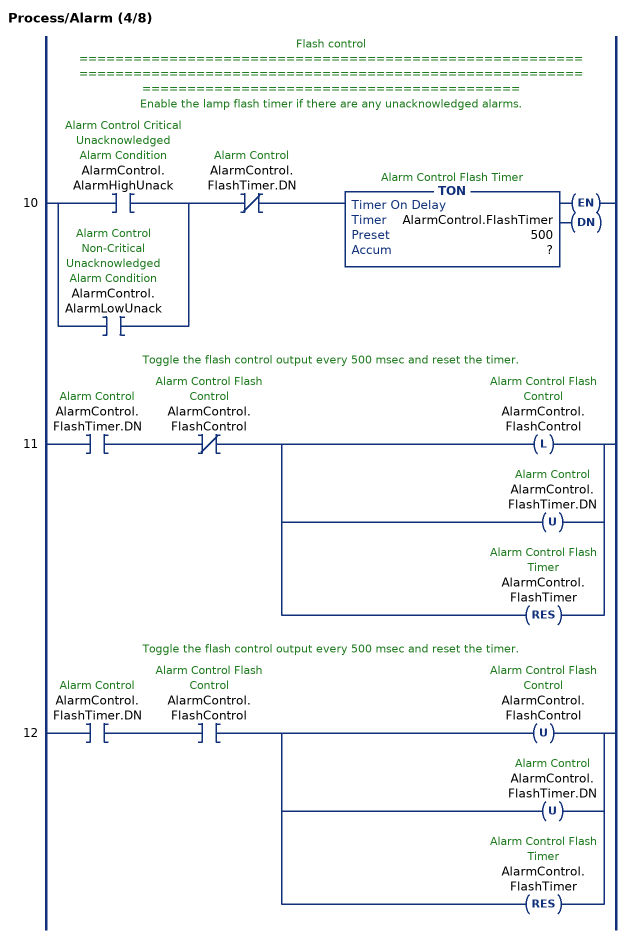
   // Flash control
   // ==========================================================================================================================================================
   // Enable the lamp flash timer if there are any unacknowledged alarms.
   10: [XIC(AlarmControl.AlarmHighUnack) ,XIC(AlarmControl.AlarmLowUnack) ]XIO(AlarmControl.FlashTimer.DN)TON(AlarmControl.FlashTimer,?,?);
   // Toggle the flash control output every 500 msec and reset the timer.
   11: XIC(AlarmControl.FlashTimer.DN)XIO(AlarmControl.FlashControl)[OTL(AlarmControl.FlashControl) ,OTU(AlarmControl.FlashTimer.DN) ,RES(AlarmControl.FlashTimer) ];
   // Toggle the flash control output every 500 msec and reset the timer.
   12: XIC(AlarmControl.FlashTimer.DN)XIC(AlarmControl.FlashControl)[OTU(AlarmControl.FlashControl) ,OTU(AlarmControl.FlashTimer.DN) ,RES(AlarmControl.FlashTimer) ];
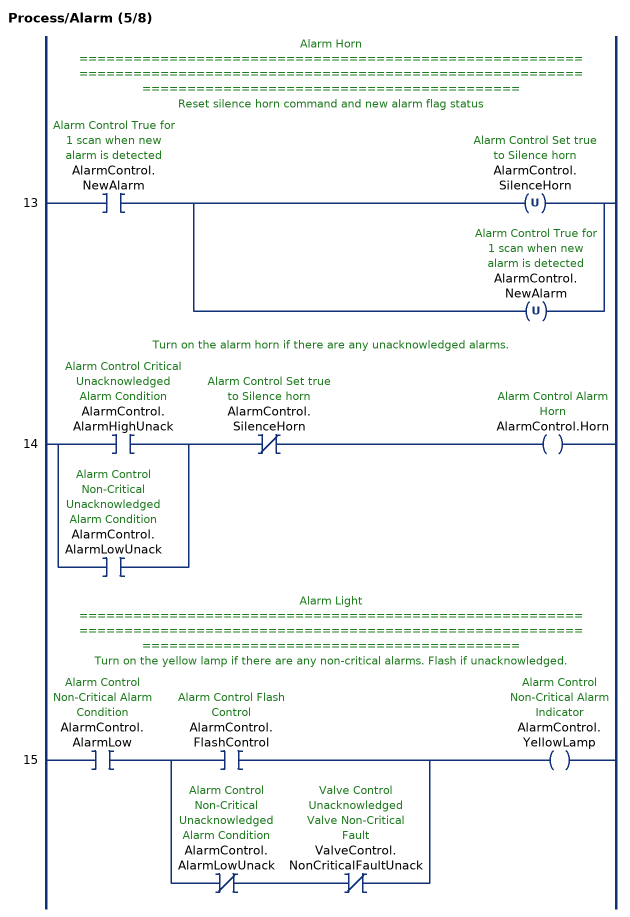
   // Alarm Horn
   // ==========================================================================================================================================================
   // Reset silence horn command and new alarm flag status
   13: XIC(AlarmControl.NewAlarm)[OTU(AlarmControl.SilenceHorn) ,OTU(AlarmControl.NewAlarm) ];
   // Turn on the alarm horn if there are any unacknowledged alarms.
   14: [XIC(AlarmControl.AlarmHighUnack) ,XIC(AlarmControl.AlarmLowUnack) ]XIO(AlarmControl.SilenceHorn)OTE(AlarmControl.Horn);
   // Alarm Light
   // ==========================================================================================================================================================
   // Turn on the yellow lamp if there are any non-critical alarms. Flash if unacknowledged.
   15: XIC(AlarmControl.AlarmLow)[XIC(AlarmControl.FlashControl) ,XIO(AlarmControl.AlarmLowUnack) XIO(ValveControl.NonCriticalFaultUnack) ]OTE(AlarmControl.YellowLamp);
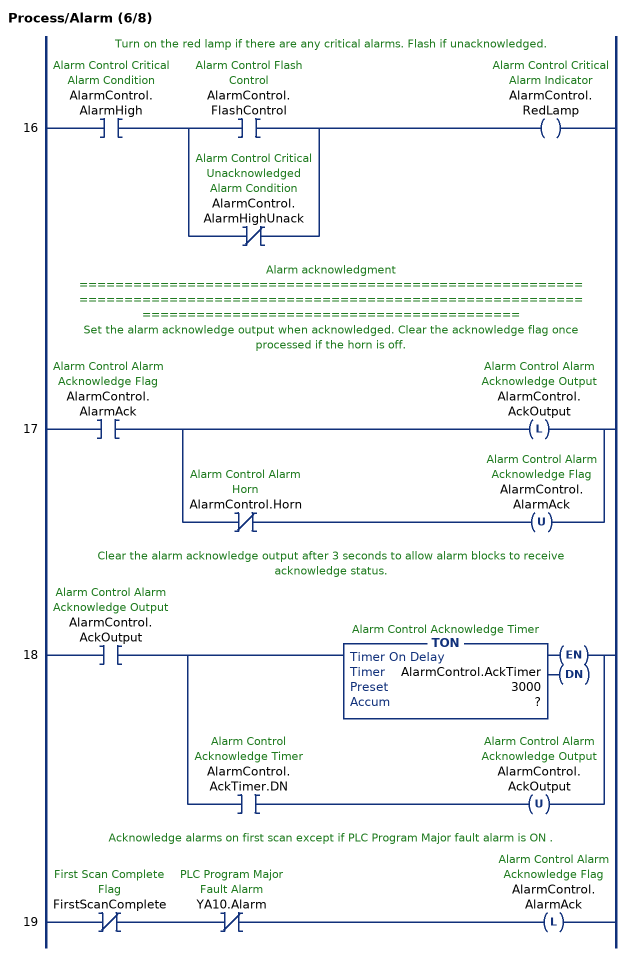
   // Turn on the red lamp if there are any critical alarms. Flash if unacknowledged.
   16: XIC(AlarmControl.AlarmHigh)[XIC(AlarmControl.FlashControl) ,XIO(AlarmControl.AlarmHighUnack) ]OTE(AlarmControl.RedLamp);
   // Alarm acknowledgment
   // ==========================================================================================================================================================
   // Set the alarm acknowledge output when acknowledged. Clear the acknowledge flag once processed if the horn is off.
   17: XIC(AlarmControl.AlarmAck)[OTL(AlarmControl.AckOutput) ,XIO(AlarmControl.Horn) OTU(AlarmControl.AlarmAck) ];
   // Clear the alarm acknowledge output after 3 seconds to allow alarm blocks to receive acknowledge status.
   18: XIC(AlarmControl.AckOutput)[TON(AlarmControl.AckTimer,?,?) ,XIC(AlarmControl.AckTimer.DN) OTU(AlarmControl.AckOutput) ];
   // Acknowledge alarms on first scan except if PLC Program Major fault alarm is ON .
   19: XIO(FirstScanComplete)XIO(YA10.Alarm)OTL(AlarmControl.AlarmAck);
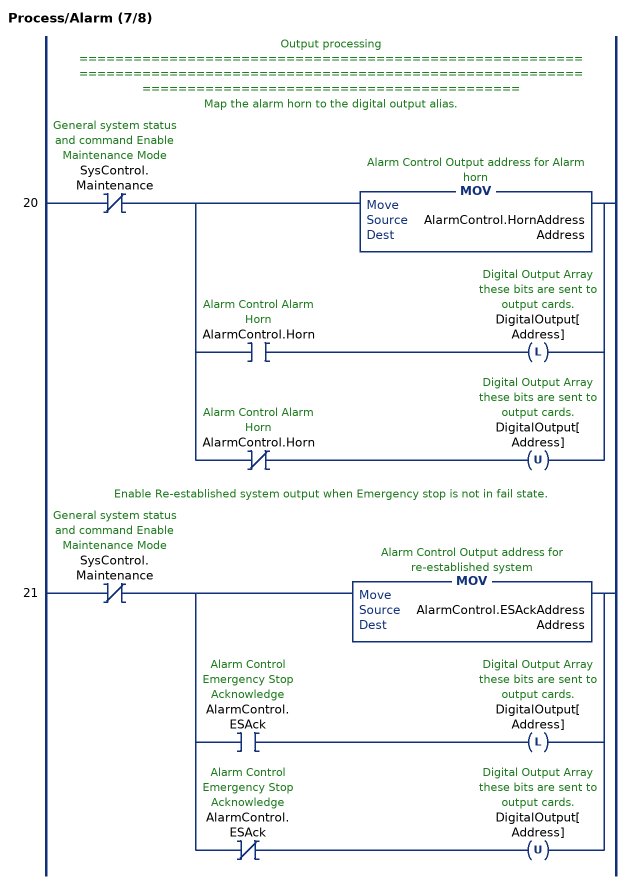
   // Output processing
   // ==========================================================================================================================================================
   // Map the alarm horn to the digital output alias.
   20: XIO(SysControl.Maintenance)[MOV(AlarmControl.HornAddress,Address) ,XIC(AlarmControl.Horn) OTL(DigitalOutput[Address]) ,XIO(AlarmControl.Horn) OTU(DigitalOutput[Address]) ];
   // Enable Re-established system output when Emergency stop is not in fail state.
   21: XIO(SysControl.Maintenance)[MOV(AlarmControl.ESAckAddress,Address) ,XIC(AlarmControl.ESAck) OTL(DigitalOutput[Address]) ,XIO(AlarmControl.ESAck) OTU(DigitalOutput[Address]) ];
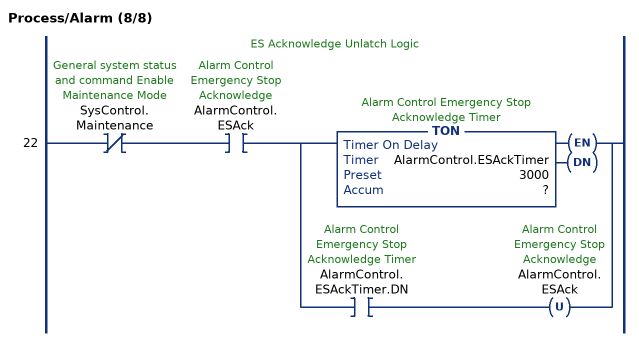
   // ES Acknowledge Unlatch Logic
   22: XIO(SysControl.Maintenance)XIC(AlarmControl.ESAck)[TON(AlarmControl.ESAckTimer,?,?) ,XIC(AlarmControl.ESAckTimer.DN) OTU(AlarmControl.ESAck) ];
END_ROUTINE
